Staubli VAL3: onShow.pgx

public program onShow()
  local num l_i
begin
  aEditItem.sComment=actdata:aActItem[nSelList].sComment
  for l_i = 0 to size(aEditItem.aActItem)-1

    aEditItem.aActItem[l_i].nIOindex=actdata:aActItem[nSelList].aActItem[l_i].nIOindex
    aEditItem.aActItem[l_i].bActive=(actdata:aActItem[nSelList].aActItem[l_i].bActive==true)
    aEditItem.aActItem[l_i].nboolValue=actdata:aActItem[nSelList].aActItem[l_i].nboolValue
    aEditItem.aActItem[l_i].nPulseValue=actdata:aActItem[nSelList].aActItem[l_i].nPulseValue
    aEditItem.aActItem[l_i].sIOtype=actdata:aActItem[nSelList].aActItem[l_i].sIOtype
    aEditItem.aActItem[l_i].sValue=actdata:aActItem[nSelList].aActItem[l_i].sValue

    sSelIO[l_i]=toString("",aEditItem.aActItem[l_i].nIOindex)
  endFor
end
